SUBAPPLICATION DummyGroup (* Platzhalter-Optionsgruppe ohne reale I/O: quittiert INIT_REQ sofort selbst per INIT_CNF (kein QI, keine Wirkung) - nuetzlich als neutraler/unbelegter Slot in einem AOption_AUI_DEMUX (z.B. fuer 'nichts ausgewaehlt' bei K=1, wenn echte Optionen erst ab K=2 beginnen) *)
  (* Standard: 61499-2; Description: Copyright (c) 2026 Meisterschulen am Ostbahnhof This program and the accompanying materials are made available under the terms of the Eclipse Public License 2.0 which is available at https://www.eclipse.org/legal/epl-2.0/ SPDX-License-Identifier: EPL-2.0 *)
  (* Version 1.0, 2026-10-13, Franz Höpfinger, Meisterschulen am Ostbahnhof, Loest das 'welcher Zahlenwert bedeutet Aus'-Problem ohne Override-Literal: ein eigener, bewusst wirkungsloser DEMUX-Slot repraesentiert den neutralen Zustand. *)
  PACKAGE MyLib_AX_Option::sys;
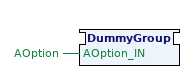
  SOCKETS
    AOption_IN : Option::AOption;
  END_SOCKETS
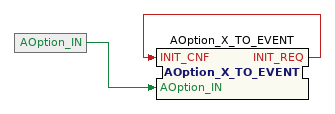
  FBS
    AOption_X_TO_EVENT : Option::conversion::AOption_X_TO_EVENT;
  END_FBS
  EVENT_CONNECTIONS
    AOption_X_TO_EVENT.INIT_REQ TO AOption_X_TO_EVENT.INIT_CNF;
  END_CONNECTIONS
  ADAPTER_CONNECTIONS
    AOption_IN TO AOption_X_TO_EVENT.AOption_IN;
  END_CONNECTIONS
END_SUBAPPLICATION
